FUNCTION_BLOCK FB 1
TITLE = Prova tedesca
VERSION : 0.1

VAR_INPUT
  Avvio : BOOL;
  Quota : ARRAY [1..3] OF INT;
END_VAR

VAR_OUTPUT
  Marcia : BOOL;
END_VAR

BEGIN
NETWORK
TITLE =
	U     E      0.0;
	UN    E      0.1;
	=     A      0.0;
	L     EW     2;
	T     MW     10;
END_FUNCTION_BLOCK
